    rq_activate_all_grippers(True)
    # end: URCap Program Node
  end
  $ 55 "zero_ftsensor()"
  zero_ftsensor()
  $ 56 "EXTT"
  $ 57 "Set GRP_3F_Enable=Off"
  set_standard_digital_out(4, False)
  $ 58 "Set BarcodeTrigger=Off"
  set_standard_digital_out(6, False)
  $ 59 "Set GRP_3F_Decap=Off"
  set_standard_digital_out(3, False)
  $ 60 "Set GRP_3F_Cap=Off"
  set_standard_digital_out(2, False)
  $ 61 "Set GRP_3F_Open=Off"
  set_standard_digital_out(5, False)
  $ 62 "PSE_T≔get_tool_free_pose(dir=[0,0,0.150], move_in_base_frame=True)"
  global PSE_T=get_tool_free_pose(dir=[0,0,0.150], move_in_base_frame=True)
  $ 63 "If is_reachable(Base_const, [PSE_T])"
  if (is_reachable(p[0.0,0.0,0.0,0.0,0.0,0.0], [PSE_T])):
    $ 64 "MoveL"
    $ 65 "PSE_T" "breakAfter"
    movel(PSE_T, a=1.2, v=0.15)
  end
  $ 677 "Thread_1"
  thread Thread_1():
    while (True):
      $ 678 "BS_Error≔IHskAndErr"
      global BS_Error=read_input_boolean_register(10)
      $ 680 "BS_Busy≔IBusy"
      global BS_Busy=read_input_boolean_register(13)
      $ 684 "BS_Complete≔ICmdExctd"
      global BS_Complete=read_input_boolean_register(12)
    end
  end
  threadId_Thread_1 = run Thread_1()
  while (True):
    $ 66 "Robot Program"
    $ 67 "MAIN"
    $ 68 "command_manager(external_control='uGO', cond_suspend=(ITM_Manipulated and AMR_AtTarget and AMR_Charging and AMR_Battery<40), cond_unsuspend=(AMR_Battery≟60))"
    command_manager(external_control="uGO", cond_suspend=(ITM_Manipulated  and  AMR_AtTarget  and  AMR_Charging  and  AMR_Battery<40), cond_unsuspend=(AMR_Battery == 60))
    $ 69 "log_state(STATE_Info)"
    log_state(STATE_Info)
    $ 70 "Switch STATE"
    switch_1 = STATE
    $ 71 "Case 1"
    if (1 == switch_1):
      $ 72 "Stopping"
      $ 73 "STATE_Info≔'Stopping'"
      global STATE_Info="Stopping"
      $ 74 "end_freedrive_mode()"
      end_freedrive_mode()
      $ 75 "Set"
      set_tcp(p[0.0,0.0,0.161,3.1415,0.0,0.0])
      $ 76 "PSE_T≔get_tool_free_pose(dir=[0,0,0.150], move_in_base_frame=True)"
      global PSE_T=get_tool_free_pose(dir=[0,0,0.150], move_in_base_frame=True)
      $ 77 "If is_reachable(Base_const, [PSE_T])"
      if (is_reachable(p[0.0,0.0,0.0,0.0,0.0,0.0], [PSE_T])):
        $ 78 "MoveL"
        $ 79 "PSE_T" "breakAfter"
        movel(PSE_T, a=1.2, v=0.15)
      end
      $ 80 "do_transition(keep_rxry=OBJ_Picked, r=0)"
      do_transition(keep_rxry=OBJ_Picked, r=0)
      $ 81 "Decapper"
      $ 82 "Set GRP_3F_Enable=Off"
      set_standard_digital_out(4, False)
      $ 83 "Set BarcodeTrigger=Off"
      set_standard_digital_out(6, False)
      $ 84 "Set GRP_3F_Decap=Off"
      set_standard_digital_out(3, False)
      $ 85 "Set GRP_3F_Cap=Off"
      set_standard_digital_out(2, False)
      $ 86 "Set GRP_3F_Open=Off"
      set_standard_digital_out(5, False)
      $ 89 "Call Sub_AMR_MiR_V3"
      Sub_AMR_MiR_V3()
      $ 90 "If stopping() and AMR_Done"
      if (stopping()  and  AMR_Done):
        $ 91 "STATE≔2"
        global STATE=2
        $ 92 "ugo_update_outputs()"
        ugo_update_outputs()
      end
    elif (2 == switch_1):
      $ 93 "Case 2"
      $ 94 "Stopped"
      $ 95 "STATE_Info≔'Stopped'"
      global STATE_Info="Stopped"
      $ 96 "Call Sub_AMR_MiR_V3"
      Sub_AMR_MiR_V3()
      $ 97 "If CMD_Reset"
      if (CMD_Reset):
        $ 98 "STATE≔3"
        global STATE=3
        $ 99 "ugo_update_outputs()"
        ugo_update_outputs()
      end
    elif (3 == switch_1):
      $ 100 "Case 3"
      $ 101 " Resetting"
      $ 102 "STATE_Info≔'Resetting'"
      global STATE_Info="Resetting"
      $ 103 "uML"
      $ 104 "reset_error()"
      reset_error()
      $ 105 "reset_warning()"
      reset_warning()
      $ 106 "PROCESS_Step≔0"
      global PROCESS_Step=0
      $ 107 "PROCESS_Info≔''"
      global PROCESS_Info=""
      $ 108 "ARM_Referenced≔ False "
      global ARM_Referenced=  False
      $ 109 "WRK_Done≔ False "
      global WRK_Done=  False
      $ 110 "ITM_Prepared≔ False "
      global ITM_Prepared=  False
      $ 111 "ITM_Manipulated≔ False "
      global ITM_Manipulated=  False
      $ 112 "STP≔0"
      global STP=0
      $ 113 "Action≔0"
      global Action=0
      $ 114 "Action_Info≔''"
      global Action_Info=""
      $ 115 "ITM_ID≔0"
      global ITM_ID=0
      $ 116 "JIG≔0"
      global JIG=0
      $ 117 "JIG_Slot≔0"
      global JIG_Slot=0
      $ 118 "Task_info≔''"
      global Task_info=""
      $ 119 "Set"
      set_tcp(p[0.0,0.0,0.161,3.1415,0.0,0.0])
      $ 120 "App"
      $ 121 "'ADD APPLICATION SPECIFIC COMMANDS'"
      # 'ADD APPLICATION SPECIFIC COMMANDS'
      $ 122 "OBJ_Type≔0"
      global OBJ_Type=0
      $ 123 "OBJ_Nbr≔0"
      global OBJ_Nbr=0
      $ 124 "If CNT_Rack_Output≥50"
      if (CNT_Rack_Output >= 50):
        $ 125 "CNT_Rack_Output≔0"
        global CNT_Rack_Output=0
      end
      $ 126 "TASK≔struct(ID=0, NAVI=struct(target=0, footprint=0, protectiveOff=0, dock=0), WORK=struct(ITM_ID_Src=0, JIG_ID_Src=0, OBJ_Nbr_Src=0, ACT_Src=0, ITM_ID_Tgt=0, JIG_ID_Tgt=0, OBJ_Nbr_Tgt=0, ACT_Tgt=0, OBJ_Type=0))"
      global TASK=struct(ID=0, NAVI=struct(target=0, footprint=0, protectiveOff=0, dock=0), WORK=struct(ITM_ID_Src=0, JIG_ID_Src=0, OBJ_Nbr_Src=0, ACT_Src=0, ITM_ID_Tgt=0, JIG_ID_Tgt=0, OBJ_Nbr_Tgt=0, ACT_Tgt=0, OBJ_Type=0))
      $ 127 "Call Sub_AMR_MiR_V3"
      Sub_AMR_MiR_V3()
      $ 128 "If resetting() and AMR_Done"
      if (resetting()  and  AMR_Done):
        $ 129 "STATE≔4"
        global STATE=4
        $ 130 "ugo_update_outputs()"
        ugo_update_outputs()
      end
    elif (4 == switch_1):
      $ 131 "Case 4"
      $ 132 "Idle"
      $ 133 "STATE_Info≔'Idle'"
      global STATE_Info="Idle"
      $ 134 "If CMD_Start"
      if (CMD_Start):
        $ 135 "STATE≔5"
        global STATE=5
        $ 136 "ugo_update_outputs()"
        ugo_update_outputs()
      end
    elif (5 == switch_1):
      $ 137 "Case 5"
      $ 138 "Starting"
      $ 139 "STATE_Info≔'Starting'"
      global STATE_Info="Starting"
      $ 140 "'ADD COMMANDS WHAT TO START WITH'"
      # 'ADD COMMANDS WHAT TO START WITH'
      $ 141 "Call Sub_AMR_MiR_V3"
      Sub_AMR_MiR_V3()
      $ 142 "get ugo data"
      $ 143 "Assign Tasks"
      $ 144 "TASK.ID = ugo_get_task()"
      TASK.ID = ugo_get_task()
      $ 145 "If TASK.ID≟1"
      if (TASK.ID == 1):
        $ 146 "Task_info≔'Charge'"
        global Task_info="Charge"
        $ 147 "Parameters"
        $ 148 "AMR_PosTarget≔1"
        global AMR_PosTarget=1
      else:
        $ 149 "ElseIf TASK.ID≟9"
        if (TASK.ID == 9):
          $ 150 "'Pick Sarstedt Rack from Variable source'"
          # 'Pick Sarstedt Rack from Variable source'
          $ 151 "Task_info≔'Navigate to Target'"
          global Task_info="Navigate to Target"
          $ 152 "Parameters"
          $ 153 "AMR_PosTarget≔UGO.read_input('00','ITM_ID')"
          global AMR_PosTarget=UGO.read_input("00","ITM_ID")
        else:
          $ 154 "ElseIf TASK.ID≟10"
          if (TASK.ID == 10):
            $ 155 "'Pick Sarstedt Rack from Variable source'"
            # 'Pick Sarstedt Rack from Variable source'
            $ 156 "Task_info≔'Pick Rack'"
            global Task_info="Pick Rack"
            $ 157 "AMR_PosTarget≔AMR_PosActual"
            global AMR_PosTarget=AMR_PosActual
            $ 158 "Parameters"
            $ 159 "ITM_ID≔UGO.read_input('00','ITM_ID')"
            global ITM_ID=UGO.read_input("00","ITM_ID")
            $ 160 "JIG≔UGO.read_input('00','JIG_ID')"
            global JIG=UGO.read_input("00","JIG_ID")
            $ 161 "OBJ_Type≔3"
            global OBJ_Type=3
          else:
            $ 163 "ElseIf TASK.ID≟11"
            if (TASK.ID == 11):
              $ 164 "'Place Sarstedt Rack on Variable target'"
              # 'Place Sarstedt Rack on Variable target'
              $ 165 "Task_info≔'Place Rack'"
              global Task_info="Place Rack"
              $ 166 "Parameters"
              $ 167 "ITM_ID≔UGO.read_input('00','ITM_ID')"
              global ITM_ID=UGO.read_input("00","ITM_ID")
              $ 168 "JIG≔UGO.read_input('00','JIG_ID')"
              global JIG=UGO.read_input("00","JIG_ID")
              $ 169 "OBJ_Type≔3"
              global OBJ_Type=3
            else:
              $ 177 "ElseIf TASK.ID≟13"
              if (TASK.ID == 13):
                $ 178 "Task_info≔'Empty racks'"
                global Task_info="Empty racks"
                $ 179 "Parameters"
                $ 180 "ITM_ID≔1"
                global ITM_ID=1
                $ 181 "AMR_PosTarget≔AMR_PosActual"
                global AMR_PosTarget=AMR_PosActual
              else:
                $ 182 "ElseIf TASK.ID≟14"
                if (TASK.ID == 14):
                  $ 183 "Task_info≔'Decap'"
                  global Task_info="Decap"
                  $ 184 "Parameters"
                  $ 185 "ITM_ID≔1"
                  global ITM_ID=1
                  $ 186 "OBJ_Type≔2"
                  global OBJ_Type=2
                  $ 187 "JIG≔7"
                  global JIG=7
                  $ 188 "AMR_PosTarget≔AMR_PosActual"
                  global AMR_PosTarget=AMR_PosActual
                else:
                  $ 189 "ElseIf TASK.ID≟99"
                  if (TASK.ID == 99):
                    $ 190 "Task_info≔'Decapping and barcode alignment'"
                    global Task_info="Decapping and barcode alignment"
                    $ 191 "Parameters"
                    $ 192 "PRC_TubNumber≔UGO.read_input('00','TubesNb')"
                    global PRC_TubNumber=UGO.read_input("00","TubesNb")
                    $ 193 "PRC_TubCounter≔0"
                    global PRC_TubCounter=0
                    $ 194 "ITM_ID≔1"
                    global ITM_ID=1
                    $ 195 "AMR_PosTarget≔AMR_PosActual"
                    global AMR_PosTarget=AMR_PosActual
                  else:
                    $ 204 "ElseIf TASK.ID≟15"
                    if (TASK.ID == 15):
                      $ 205 "Task_info≔'Unoad Centrifuge'"
                      global Task_info="Unoad Centrifuge"
                      $ 206 "Parameters"
                      $ 207 "PRC_RackCounter≔0"
                      global PRC_RackCounter=0
                      $ 208 "TASK.WORK.ITM_ID_Src=2"
                      TASK.WORK.ITM_ID_Src=2
                      $ 209 "TASK.WORK.ITM_ID_Tgt=1"
                      TASK.WORK.ITM_ID_Tgt=1
                      $ 210 "AMR_PosTarget≔4"
                      global AMR_PosTarget=4
                      $ 211 "AMR_FootprintID≔1"
                      global AMR_FootprintID=1
                    else:
                      $ 230 "Else" "noBreak"
                      $ 231 "set_error(ERROR_WRONG_ORDER)"
                      set_error(ERROR_WRONG_ORDER)
                    end
                  end
                end
              end
            end
          end
        end
      end
      $ 232 "test ugo"
      $ 233 "Wait: 0.2"
      sleep(0.2)
      $ 234 "ugo_update_outputs()"
      ugo_update_outputs()
      $ 235 "If starting() and AMR_Done"
      if (starting()  and  AMR_Done):
        $ 236 "log_message(Task_info, 'New Task: ')"
        log_message(Task_info, "New Task: ")
        $ 237 "log_message(to_str(TASK.ID), 'Task_ID: ')"
        log_message(to_str(TASK.ID), "Task_ID: ")
        $ 238 "do_transition(keep_rxry=OBJ_Picked)"
        do_transition(keep_rxry=OBJ_Picked)
        $ 239 "STATE≔6"
        global STATE=6
        $ 240 "ugo_update_outputs()"
        ugo_update_outputs()
      end
    elif (6 == switch_1):
      $ 241 "Case 6"
      $ 242 "Execute"
      $ 243 "STATE_Info≔'Execute'"
      global STATE_Info="Execute"
      $ 244 "If  not CMD_Hold and not CMD_Suspend"
      global thread_flag_244=0
      thread Thread_if_244():
        $ 245 "Switch PROCESS_Step"
        switch_2 = PROCESS_Step
        $ 246 "Case 0"
        if (0 == switch_2):
          $ 247 "PROCESS_Info≔'process control'"
          global PROCESS_Info="process control"
          $ 248 "log_process(PROCESS_Info)"
          log_process(PROCESS_Info)
          $ 249 "process control"
          $ 250 "If  not AMR_AtTarget"
          if (  not  AMR_AtTarget):
            $ 251 "PROCESS_Step≔1"
            global PROCESS_Step=1
          else:
            $ 252 "ElseIf (( not ITM_Prepared and  not WRK_Done) or (ITM_Prepared and WRK_Done))"
            if (((  not  ITM_Prepared  and    not  WRK_Done)  or  (ITM_Prepared  and  WRK_Done))):
              $ 253 "PROCESS_Step≔2"
              global PROCESS_Step=2
            else:
              $ 254 "ElseIf  not WRK_Done"
              if (  not  WRK_Done):
                $ 255 "PROCESS_Step≔3"
                global PROCESS_Step=3
              else:
                $ 256 "Else" "noBreak"
                $ 257 "task finished"
                $ 258 "PROCESS_Info≔''"
                global PROCESS_Info=""
                $ 259 "STATE≔7"
                global STATE=7
                $ 260 "ugo_update_outputs()"
                ugo_update_outputs()
              end
            end
          end
        elif (1 == switch_2):
          $ 261 "Case 1"
          $ 262 "navigate"
          $ 263 "'MOVING THE uML'"
          # 'MOVING THE uML'
          $ 264 "PROCESS_Info≔'move to target'"
          global PROCESS_Info="move to target"
          $ 265 "log_process(PROCESS_Info)"
          log_process(PROCESS_Info)
          $ 266 "If TASK.ID≟1"
          if (TASK.ID == 1):
            $ 267 "Action≔51"
            global Action=51
          else:
            $ 268 "Else" "noBreak"
            $ 269 "Action≔52"
            global Action=52
          end
          $ 270 "Call Sub_AMR_MiR_V3"
          Sub_AMR_MiR_V3()
          $ 271 "If AMR_Done"
          if (AMR_Done):
            $ 272 "PROCESS_Step≔0"
            global PROCESS_Step=0
          end
        elif (2 == switch_2):
          $ 273 "Case 2"
          $ 274 "prepare"
          $ 275 "'THINGS THAT HAVE TO BE DONE ONCE IN A SEQUENCE,WORKFLOW'"
          # 'THINGS THAT HAVE TO BE DONE ONCE IN A SEQUENCE,WORKFLOW'
          $ 276 "PROCESS_Info≔'prepare for work'"
          global PROCESS_Info="prepare for work"
          $ 277 "log_process(PROCESS_Info)"
          log_process(PROCESS_Info)
          $ 278 "If TASK.WORK.ITM_ID_Src>1"
          if (TASK.WORK.ITM_ID_Src>1):
            $ 279 "ITM_ID≔TASK.WORK.ITM_ID_Src"
            global ITM_ID=TASK.WORK.ITM_ID_Src
          else:
            $ 280 "ElseIf TASK.WORK.ITM_ID_Tgt>1"
            if (TASK.WORK.ITM_ID_Tgt>1):
              $ 281 "ITM_ID≔TASK.WORK.ITM_ID_Tgt"
              global ITM_ID=TASK.WORK.ITM_ID_Tgt
            end
          end
          $ 282 "If  not ARM_Referenced and (ITM_ID≠0)"
          if (  not  ARM_Referenced  and  (ITM_ID != 0)):
            $ 283 "STP≔1"
            global STP=1
          else:
            $ 284 "ElseIf ARM_Referenced or (ITM_ID≟0)"
            if (ARM_Referenced  or  (ITM_ID == 0)):
              $ 285 "STP≔2"
              global STP=2
            end
          end
          $ 286 "Switch STP"
          switch_3 = STP
          $ 287 "Case 1"
          if (1 == switch_3):
            $ 288 "reference"
            $ 289 "STP_Info≔'reference at target position'"
            global STP_Info="reference at target position"
            $ 290 "log_step(STP_Info)"
            log_step(STP_Info)
            $ 291 "If ITM_ID≟1"
            if (ITM_ID == 1):
              $ 292 "CAM_Done≔ True "
              global CAM_Done=  True
            else:
              $ 293 "Else" "noBreak"
              $ 294 "Action≔131"
              global Action=131
              $ 295 "Call Sub_Vision_V18"
              Sub_Vision_V18()
            end
            $ 297 "If CAM_Done and  not ERROR.FLAG"
            if (CAM_Done  and    not  ERROR.FLAG):
              $ 298 "log_step('ARM referenced')"
              log_step("ARM referenced")
              $ 299 "ARM_Referenced≔ True "
              global ARM_Referenced=  True
            end
          elif (2 == switch_3):
            $ 300 "Case 2"
            $ 301 "manipulate"
            $ 302 "STP_Info≔'manipulate item'"
            global STP_Info="manipulate item"
            $ 303 "log_step(STP_Info)"
            log_step(STP_Info)
            $ 304 "'In case pressing button is needed'"
            # 'In case pressing button is needed'
            $ 305 "If found_in_list(ITM_ID, ITM_ID_List)"
            if (found_in_list(ITM_ID, ITM_ID_List)):
              $ 306 "Switch ITM_ID"
              switch_4 = ITM_ID
              $ 307 "Case 0"
              if (0 == switch_4):
                $ 308 "ITM_Manipulated≔ not ITM_Manipulated"
                global ITM_Manipulated=  not  ITM_Manipulated
              elif (1 == switch_4):
                $ 309 "Case 1"
                $ 310 "ITM_Manipulated≔ not ITM_Manipulated"
                global ITM_Manipulated=  not  ITM_Manipulated
              elif (2 == switch_4):
                $ 311 "Case 2"
              else:
                $ 321 "Default Case"
                $ 322 "ITM_Manipulated≔ not ITM_Manipulated"
                global ITM_Manipulated=  not  ITM_Manipulated
              end
            end
          end
          $ 323 "ITM_Prepared≔(ITM_Manipulated or  not found_in_list(ITM_ID, ITM_ID_List)) and (ARM_Referenced or ITM_ID≟0) and  not WRK_Done"
          global ITM_Prepared=(ITM_Manipulated  or    not  found_in_list(ITM_ID, ITM_ID_List))  and  (ARM_Referenced  or  ITM_ID == 0)  and    not  WRK_Done
          $ 324 "STP≔0"
          global STP=0
          $ 325 "STP_Info≔''"
          global STP_Info=""
          $ 326 "PROCESS_Step≔0"
          global PROCESS_Step=0
        elif (3 == switch_2):
          $ 327 "Case 3"
          $ 328 "work"
          $ 329 "'ADD EVERY MACHINE, OBJECT, STATION TO WORK ON'"
          # 'ADD EVERY MACHINE, OBJECT, STATION TO WORK ON'
          $ 330 "Switch ITM_ID"
          switch_3 = ITM_ID
          $ 331 "Case 1"
          if (1 == switch_3):
            $ 332 "uLM"
            $ 333 "If TASK.ID≟12"
            if (TASK.ID == 12):
              $ 334 "fill racks"
              $ 335 "Action≔151"
              global Action=151
              $ 336 "Call Sub_Vision_V18"
              Sub_Vision_V18()
              $ 337 "If  not ERROR.FLAG"
              if (  not  ERROR.FLAG):
                $ 338 "Actions for the task"
                $ 339 "Action≔1"
                global Action=1
                $ 340 "JIG≔2"
                global JIG=2
                $ 341 "JIG_Slot≔CAM_Result[0]"
                global JIG_Slot=CAM_Result[0]
                $ 342 "OBJ_Nbr≔CAM_Result[0]"
                global OBJ_Nbr=CAM_Result[0]
                $ 343 "OBJ_Type≔2"
                global OBJ_Type=2
                $ 344 "Call Sub_Action_V4"
                Sub_Action_V4()
                $ 345 "If OBJ_Picked"
                if (OBJ_Picked):
                  $ 346 "CAM_Result.remove(0)"
                  CAM_Result.remove(0)
                  $ 347 "PRC_TubCounter≔PRC_TubCounter+1"
                  global PRC_TubCounter=PRC_TubCounter+1
                  $ 348 "If PRC_TubCounter%4≟0"
                  if (PRC_TubCounter%4 == 0):
                    $ 349 "JIG_Slot≔4"
                    global JIG_Slot=4
                  else:
                    $ 350 "Else" "noBreak"
                    $ 351 "JIG_Slot≔PRC_TubCounter%4"
                    global JIG_Slot=PRC_TubCounter%4
                  end
                  $ 352 "OBJ_Nbr≔ceil(PRC_TubCounter/4)"
                  global OBJ_Nbr=ceil(PRC_TubCounter/4)
                  $ 353 "Action≔2"
                  global Action=2
                  $ 354 "JIG≔4"
                  global JIG=4
                  $ 355 "Call Sub_Action_V4"
                  Sub_Action_V4()
                  $ 356 "Action≔151"
                  global Action=151
                  $ 357 "Call Sub_Vision_V18"
                  Sub_Vision_V18()
                end
              end
              $ 358 "If (CAM_Captures≥CAM_PRM_Retries) or (PRC_TubCounter≥32)"
              if ((CAM_Captures >= CAM_PRM_Retries)  or  (PRC_TubCounter >= 32)):
                $ 359 "PROCESS_Step≔0"
                global PROCESS_Step=0
                $ 360 "WRK_Done≔ True "
                global WRK_Done=  True
              end
            else:
              $ 364 "ElseIf TASK.ID≟10"
              if (TASK.ID == 10):
                $ 365 "Pick Rack"
                $ 366 "Action≔131"
                global Action=131
                $ 367 "Call Sub_Vision_V18"
                Sub_Vision_V18()
                $ 368 "Action≔1"
                global Action=1
                $ 369 "Call Sub_Action_V4"
                Sub_Action_V4()
                $ 370 "PROCESS_Step≔0"
                global PROCESS_Step=0
                $ 371 "WRK_Done≔ True "
                global WRK_Done=  True
              else:
                $ 372 "ElseIf TASK.ID≟11"
                if (TASK.ID == 11):
                  $ 373 "Place Rack"
                  $ 374 "Action≔2"
                  global Action=2
                  $ 375 "Call Sub_Action_V4"
                  Sub_Action_V4()
                  $ 376 "PROCESS_Step≔0"
                  global PROCESS_Step=0
                  $ 377 "WRK_Done≔ True "
                  global WRK_Done=  True
                else:
                  $ 378 "ElseIf TASK.ID≟13"
                  if (TASK.ID == 13):
                    $ 379 "empty racks"
                    $ 380 "pick"
                    $ 381 "Action≔1"
                    global Action=1
                    $ 382 "JIG≔4"
                    global JIG=4
                    $ 383 "If PRC_TubCounter%4≟0"
                    if (PRC_TubCounter%4 == 0):
                      $ 384 "JIG_Slot≔4"
                      global JIG_Slot=4
                    else:
                      $ 385 "Else" "noBreak"
                      $ 386 "JIG_Slot≔PRC_TubCounter%4"
                      global JIG_Slot=PRC_TubCounter%4
                    end
                    $ 387 "OBJ_Nbr≔ceil(PRC_TubCounter/4)"
                    global OBJ_Nbr=ceil(PRC_TubCounter/4)
                    $ 388 "OBJ_Type≔2"
                    global OBJ_Type=2
                    $ 389 "Call Sub_Action_V4"
                    Sub_Action_V4()
                    $ 390 "If OBJ_Picked"
                    if (OBJ_Picked):
                      $ 391 "Action≔2"
                      global Action=2
                      $ 392 "JIG≔3"
                      global JIG=3
                      $ 393 "JIG_Slot≔1"
                      global JIG_Slot=1
                      $ 394 "CNT_Rack_Output≔CNT_Rack_Output + 1"
                      global CNT_Rack_Output=CNT_Rack_Output + 1
                      $ 395 "OBJ_Nbr≔CNT_Rack_Output"
                      global OBJ_Nbr=CNT_Rack_Output
                      $ 396 "Call Sub_Action_V4"
                      Sub_Action_V4()
                      $ 397 "If  not ERROR.FLAG"
                      if (  not  ERROR.FLAG):
                        $ 398 "PRC_TubCounter≔PRC_TubCounter - 1"
                        global PRC_TubCounter=PRC_TubCounter - 1
                      end
                    end
                    $ 399 "If CNT_Rack_Output≥50 or PRC_TubCounter≤0"
                    if (CNT_Rack_Output >= 50  or  PRC_TubCounter <= 0):
                      $ 400 "PROCESS_Step≔0"
                      global PROCESS_Step=0
                      $ 401 "WRK_Done≔ True "
                      global WRK_Done=  True
                    end
                  else:
                    $ 402 "ElseIf TASK.ID≟14"
                    if (TASK.ID == 14):
                      $ 405 "samples≔ True "
                      global samples=  True
                      $ 406 "Loop samples≟ True "
                      while (samples ==   True  ):
                        $ 412 "JIG≔1"
                        global JIG=1
                        $ 413 "Action≔11"
                        global Action=11
                        $ 414 "Call Sub_Action_V4"
                        Sub_Action_V4()
                        $ 415 "Action≔12"
                        global Action=12
                        $ 416 "Call Sub_Action_V4"
                        Sub_Action_V4()
                        $ 417 "Action≔2"
                        global Action=2
                        $ 418 "JIG≔6"
                        global JIG=6
                        $ 419 "Call Sub_Action_V4"
                        Sub_Action_V4()
                        $ 420 "Action≔13"
                        global Action=13
                        $ 421 "Call Sub_Action_V4"
                        Sub_Action_V4()
                        $ 422 "Action≔1"
                        global Action=1
                        $ 423 "JIG≔1"
                        global JIG=1
                        $ 424 "Call Sub_Action_V4"
                        Sub_Action_V4()
                      end
                    end
                  end
                end
              end
            end
          elif (2 == switch_3):
            $ 428 "Case 2"
          elif (20 == switch_3):
            $ 470 "Case 20"
          else:
            $ 532 "Default Case"
            $ 533 "WRK_Done≔ True "
            global WRK_Done=  True
            $ 534 "PROCESS_Step≔0"
            global PROCESS_Step=0
          end
        end
        thread_flag_244 = 1
      end
      if (  not  CMD_Hold and not CMD_Suspend):
        global thread_handler_244=run Thread_if_244()
        while (thread_flag_244 == 0):
          if not(  not  CMD_Hold and not CMD_Suspend):
            kill thread_handler_244
            thread_flag_244 = 2
          else:
            sync()
          end
        end
      else:
        thread_flag_244 = 2
      end
      $ 535 "If CMD_Hold"
      if (CMD_Hold):
        $ 536 "STATE≔9"
        global STATE=9
        $ 537 "ugo_update_outputs()"
        ugo_update_outputs()
      else:
        $ 538 "ElseIf CMD_Suspend"
        if (CMD_Suspend):
          $ 539 "STATE≔12"
          global STATE=12
          $ 540 "ugo_update_outputs()"
          ugo_update_outputs()
        end
      end
    elif (7 == switch_1):
      $ 541 "Case 7"
      $ 542 "Completing"
      $ 543 "STATE_Info≔'Completing'"
      global STATE_Info="Completing"
      $ 544 "'ADD COMMANDS FOR COMPLETING THE PROCESS'"
      # 'ADD COMMANDS FOR COMPLETING THE PROCESS'
      $ 545 "do_transition(keep_rxry=OBJ_Picked)"
      do_transition(keep_rxry=OBJ_Picked)
      $ 546 "Call Sub_AMR_MiR_V3"
      Sub_AMR_MiR_V3()
      $ 547 "If completing() and AMR_Done"
      if (completing()  and  AMR_Done):
        $ 548 "STATE≔8"
        global STATE=8
        $ 549 "ugo_update_outputs()"
        ugo_update_outputs()
      end
    elif (8 == switch_1):
      $ 550 "Case 8"
      $ 551 "Complete"
      $ 552 "STATE_Info≔'Complete'"
      global STATE_Info="Complete"
      $ 553 "If CMD_Reset"
      if (CMD_Reset):
        $ 554 "STATE≔3"
        global STATE=3
        $ 555 "ugo_update_outputs()"
        ugo_update_outputs()
      end
    elif (9 == switch_1):
      $ 556 "Case 9"
      $ 557 "Holding"
      $ 558 "STATE_Info≔'Holding'"
      global STATE_Info="Holding"
      $ 559 "stopl(0.5)"
      stopl(0.5)
      $ 560 "Call Sub_AMR_MiR_V3"
      Sub_AMR_MiR_V3()
      $ 561 "If holding() and AMR_Done"
      if (holding()  and  AMR_Done):
        $ 562 "STATE≔10"
        global STATE=10
        $ 563 "ugo_update_outputs()"
        ugo_update_outputs()
      end
    elif (10 == switch_1):
      $ 564 "Case 10"
      $ 565 "Held"
      $ 566 "STATE_Info≔'Held'"
      global STATE_Info="Held"
      $ 567 "If CMD_Unhold"
      if (CMD_Unhold):
        $ 568 "end_freedrive_mode()"
        end_freedrive_mode()
        $ 569 "STATE≔11"
        global STATE=11
        $ 570 "ugo_update_outputs()"
        ugo_update_outputs()
      else:
        $ 571 "ElseIf FNC_Freedrive"
        if (FNC_Freedrive):
          $ 572 "freedrive_mode()"
          freedrive_mode()
        else:
          $ 573 "Else" "noBreak"
          $ 574 "end_freedrive_mode()"
          end_freedrive_mode()
        end
      end
    elif (11 == switch_1):
      $ 575 "Case 11"
      $ 576 "Unholding"
      $ 577 "STATE_Info≔'Unholding'"
      global STATE_Info="Unholding"
      $ 578 "Clearing"
      $ 579 "Switch ERROR.ID"
      switch_2 = ERROR.ID
      $ 580 "Case 1002"
      if (1002 == switch_2):
        $ 581 "AMR_AtTarget≔ False "
        global AMR_AtTarget=  False
        $ 582 "ARM_Referenced≔ False "
        global ARM_Referenced=  False
        $ 583 "ITM_Prepared≔ False "
        global ITM_Prepared=  False
        $ 584 "PROCESS_Step≔1"
        global PROCESS_Step=1
      elif (2007 == switch_2):
        $ 585 "Case 2007"
        $ 586 "PROCESS_Step≔1"
        global PROCESS_Step=1
      end
      $ 587 "reset_error()"
      reset_error()
      $ 588 "reset_warning()"
      reset_warning()
      $ 589 "OBJ_Picked≔gripper_has_object()"
      global OBJ_Picked=gripper_has_object()
      $ 590 "Call Sub_AMR_MiR_V3"
      Sub_AMR_MiR_V3()
      $ 591 "If unholding() and AMR_Done"
      if (unholding()  and  AMR_Done):
        $ 592 "STATE≔6"
        global STATE=6
        $ 593 "ugo_update_outputs()"
        ugo_update_outputs()
      end
    elif (12 == switch_1):
      $ 594 "Case 12"
      $ 595 "Suspending"
      $ 596 "STATE_Info≔'Suspending'"
      global STATE_Info="Suspending"
      $ 597 "PROCESS_Info≔str_cat(PROCESS_Info, ' suspended')"
      global PROCESS_Info=str_cat(PROCESS_Info, " suspended")
      $ 598 "If suspending()"
      if (suspending()):
        $ 599 "STATE≔13"
        global STATE=13
        $ 600 "ugo_update_outputs()"
        ugo_update_outputs()
      end
    elif (13 == switch_1):
      $ 601 "Case 13"
      $ 602 "Suspended"
      $ 603 "STATE_Info≔'Suspended'"
      global STATE_Info="Suspended"
      $ 604 "Call Sub_AMR_MiR_V3"
      Sub_AMR_MiR_V3()
      $ 605 "If CMD_Unsuspend"
      if (CMD_Unsuspend):
        $ 606 "STATE≔14"
        global STATE=14
        $ 607 "ugo_update_outputs()"
        ugo_update_outputs()
      end
    elif (14 == switch_1):
      $ 608 "Case 14"
      $ 609 "Unsuspending"
      $ 610 "STATE_Info≔'Unsuspending'"
      global STATE_Info="Unsuspending"
      $ 611 "PROCESS_Step≔0"
      global PROCESS_Step=0
      $ 612 "If unsuspending()"
      if (unsuspending()):
        $ 613 "STATE≔6"
        global STATE=6
        $ 614 "ugo_update_outputs()"
        ugo_update_outputs()
      end
    elif (15 == switch_1):
      $ 615 "Case 15"
      $ 616 "Aborting"
      $ 617 "STATE_Info≔'Aborting'"
      global STATE_Info="Aborting"
      $ 618 "If aborting()"
      if (aborting()):
        $ 619 "STATE≔16"
        global STATE=16
        $ 620 "ugo_update_outputs()"
        ugo_update_outputs()
      end
    elif (16 == switch_1):
      $ 621 "Case 16"
      $ 622 "Aborted"
      $ 623 "STATE_Info≔'Aborted'"
      global STATE_Info="Aborted"
      $ 624 "If CMD_Clear"
      if (CMD_Clear):
        $ 625 "STATE≔17"
        global STATE=17
        $ 626 "ugo_update_outputs()"
        ugo_update_outputs()
      end
    elif (17 == switch_1):
      $ 627 "Case 17"
      $ 628 "Clearing"
      $ 629 "STATE_Info≔'Clearing'"
      global STATE_Info="Clearing"
      $ 630 "Clearing"
      $ 631 "reset_warning()"
      reset_warning()
      $ 632 "reset_error()"
      reset_error()
      $ 633 "If clearing()"
      if (clearing()):
        $ 634 "STATE≔2"
        global STATE=2
        $ 635 "ugo_update_outputs()"
        ugo_update_outputs()
      end
    end
    $ 636 "log_state(STATE_Info)"
    log_state(STATE_Info)
    $ 637 "log_warning(WARNING.MSG)"
    log_warning(WARNING.MSG)
    $ 638 "log_error(ERROR.MSG)"
    log_error(ERROR.MSG)
    $ 639 "Times"
    $ 640 "Switch STATE"
    switch_1 = STATE
    $ 641 "Case 1"
    if (1 == switch_1):
      $ 642 "TM_St_Stopping≔get_time(STATE_Times[STATE-1])"
      global TM_St_Stopping=get_time(STATE_Times[STATE-1])
    elif (2 == switch_1):
      $ 643 "Case 2"
      $ 644 "TM_St_Stopped≔get_time(STATE_Times[STATE-1])"
      global TM_St_Stopped=get_time(STATE_Times[STATE-1])
    elif (3 == switch_1):
      $ 645 "Case 3"
      $ 646 "TM_St_Resetting≔get_time(STATE_Times[STATE-1])"
      global TM_St_Resetting=get_time(STATE_Times[STATE-1])
    elif (4 == switch_1):
      $ 647 "Case 4"
      $ 648 "TM_St_Idle≔get_time(STATE_Times[STATE-1])"
      global TM_St_Idle=get_time(STATE_Times[STATE-1])
    elif (5 == switch_1):
      $ 649 "Case 5"
      $ 650 "TM_St_Starting≔get_time(STATE_Times[STATE-1])"
      global TM_St_Starting=get_time(STATE_Times[STATE-1])
    elif (6 == switch_1):
      $ 651 "Case 6"
      $ 652 "TM_St_Execute≔get_time(STATE_Times[STATE-1])"
      global TM_St_Execute=get_time(STATE_Times[STATE-1])
    elif (7 == switch_1):
      $ 653 "Case 7"
      $ 654 "TM_St_Completin≔get_time(STATE_Times[STATE-1])"
      global TM_St_Completin=get_time(STATE_Times[STATE-1])
    elif (8 == switch_1):
      $ 655 "Case 8"
      $ 656 "TM_St_Complete≔get_time(STATE_Times[STATE-1])"
      global TM_St_Complete=get_time(STATE_Times[STATE-1])
    elif (9 == switch_1):
      $ 657 "Case 9"
      $ 658 "TM_St_Holding≔get_time(STATE_Times[STATE-1])"
      global TM_St_Holding=get_time(STATE_Times[STATE-1])
    elif (10 == switch_1):
      $ 659 "Case 10"
      $ 660 "TM_St_Held≔get_time(STATE_Times[STATE-1])"
      global TM_St_Held=get_time(STATE_Times[STATE-1])
    elif (11 == switch_1):
      $ 661 "Case 11"
      $ 662 "TM_St_Unholding≔get_time(STATE_Times[STATE-1])"
      global TM_St_Unholding=get_time(STATE_Times[STATE-1])
    elif (12 == switch_1):
      $ 663 "Case 12"
      $ 664 "TM_St_Suspendin≔get_time(STATE_Times[STATE-1])"
      global TM_St_Suspendin=get_time(STATE_Times[STATE-1])
    elif (13 == switch_1):
      $ 665 "Case 13"
      $ 666 "TM_St_Suspended≔get_time(STATE_Times[STATE-1])"
      global TM_St_Suspended=get_time(STATE_Times[STATE-1])
    elif (14 == switch_1):
      $ 667 "Case 14"
      $ 668 "TM_St_Unsuspend≔get_time(STATE_Times[STATE-1])"
      global TM_St_Unsuspend=get_time(STATE_Times[STATE-1])
    elif (15 == switch_1):
      $ 669 "Case 15"
      $ 670 "TM_St_Aborting≔get_time(STATE_Times[STATE-1])"
      global TM_St_Aborting=get_time(STATE_Times[STATE-1])
    elif (16 == switch_1):
      $ 671 "Case 16"
      $ 672 "TM_St_Aborted≔get_time(STATE_Times[STATE-1])"
      global TM_St_Aborted=get_time(STATE_Times[STATE-1])
    elif (17 == switch_1):
      $ 673 "Case 17"
      $ 674 "TM_St_Clearing≔get_time(STATE_Times[STATE-1])"
      global TM_St_Clearing=get_time(STATE_Times[STATE-1])
    end
    $ 676 "Wait: 0.1"
    sleep(0.1)
  end
end
